FUNCTION_BLOCK Agua_Reuso (* Agua de reuso (serie 1000) - HidrycoLib *)
  (* Standard: 61499-2 *)
  (* Version 1.3, 20/10/2026, Hidryco, Hidryco, 1.3: simbolo sBoiaL (boia animada, verde/vermelho/cinza sem comunicacao). 1.2: o MGE do PCM Agua Reuso (MGE_1000) sai do CAT: passa a ser a instancia MGE_AGUA_REUSO do frame de MGEs do ETE_TJ; saem as saidas e tags do MGE. 1.1: MGE_1000 passa a ser o MGE_Generico (PM5300 pelo HW CAT PM53xxMbtcp, falta de fase e H/L de tensao e corrente); saidas stsFaltaFaseMGE, stsAlarmeMGE e stsPotenciaAtivaMGE; sai o cfgMonitoraMGE e o symlink stsConexaoMGE. 1.0: agua de reuso (serie 1000), so monitoracao. 1000-PIT-01/02 (Sensor_Generico, 4-20 mA, nivel) pelos symlinks ${PATH}PIT_1000_0x.stsSensorBruto; boia 1000-LSL-01 por ${PATH}stsBoiaLSL; comunicacao por ${PATH}stsFalhaRemota1 (BOOL, cartao), ${PATH}stsConexaoRemota2 e ${PATH}stsConexaoMGE (INT, connStatusInt); MGE do PCM Agua Reuso no MGE_1000. Valores e alarmes nas saidas do CAT. *)
  PACKAGE Hidryco.HidrycoLib;
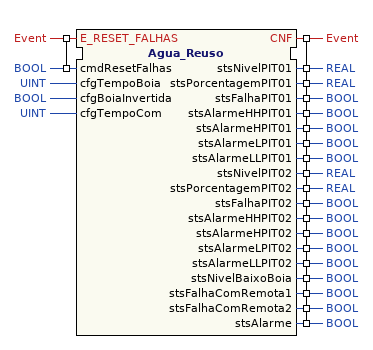
  EVENT_INPUT
    E_RESET_FALHAS WITH cmdResetFalhas; (* Reset pelo processo (sensores) com cmdResetFalhas = TRUE *)
  END_EVENT
  EVENT_OUTPUT
    CNF WITH stsNivelPIT01, stsPorcentagemPIT01, stsFalhaPIT01, stsAlarmeHHPIT01, stsAlarmeHPIT01, stsAlarmeLPIT01, stsAlarmeLLPIT01, stsNivelPIT02, stsPorcentagemPIT02, stsFalhaPIT02, stsAlarmeHHPIT02, stsAlarmeHPIT02, stsAlarmeLPIT02, stsAlarmeLLPIT02, stsNivelBaixoBoia, stsFalhaComRemota1, stsFalhaComRemota2, stsAlarme; (* Valores e alarmes (so na mudanca) *)
  END_EVENT
  VAR_INPUT
    cmdResetFalhas : BOOL; (* TRUE = reset (com o evento E_RESET_FALHAS) *)
    cfgTempoBoia : UINT := 10; (* Tempo (s) da boia 1000-LSL-01 abaixada para confirmar o nivel baixo *)
    cfgBoiaInvertida : BOOL := FALSE; (* FALSE: entrada da boia TRUE = nivel normal (boia levantada). TRUE: entrada TRUE = nivel baixo *)
    cfgTempoCom : UINT := 5; (* Tempo (s) sem comunicacao para confirmar a falha das remotas *)
  END_VAR
  VAR_OUTPUT
    stsNivelPIT01 : REAL; (* Nivel PIT_1000_01 (unidade de engenharia do sensor; 0 com o sinal em falha) *)
    stsPorcentagemPIT01 : REAL; (* Nivel PIT_1000_01 em % da altura maxima *)
    stsFalhaPIT01 : BOOL; (* Falha do sensor PIT_1000_01 (memorizada ate o reset) *)
    stsAlarmeHHPIT01 : BOOL; (* Alarme HH do PIT_1000_01 *)
    stsAlarmeHPIT01 : BOOL; (* Alarme H do PIT_1000_01 *)
    stsAlarmeLPIT01 : BOOL; (* Alarme L do PIT_1000_01 *)
    stsAlarmeLLPIT01 : BOOL; (* Alarme LL do PIT_1000_01 *)
    stsNivelPIT02 : REAL; (* Nivel PIT_1000_02 (unidade de engenharia do sensor; 0 com o sinal em falha) *)
    stsPorcentagemPIT02 : REAL; (* Nivel PIT_1000_02 em % da altura maxima *)
    stsFalhaPIT02 : BOOL; (* Falha do sensor PIT_1000_02 (memorizada ate o reset) *)
    stsAlarmeHHPIT02 : BOOL; (* Alarme HH do PIT_1000_02 *)
    stsAlarmeHPIT02 : BOOL; (* Alarme H do PIT_1000_02 *)
    stsAlarmeLPIT02 : BOOL; (* Alarme L do PIT_1000_02 *)
    stsAlarmeLLPIT02 : BOOL; (* Alarme LL do PIT_1000_02 *)
    stsNivelBaixoBoia : BOOL; (* Nivel baixo pela boia 1000-LSL-01 (confirmado por cfgTempoBoia) *)
    stsFalhaComRemota1 : BOOL; (* Falha de comunicacao com a remota 1 da Subestacao (boia) *)
    stsFalhaComRemota2 : BOOL; (* Falha de comunicacao com a remota 2 da Subestacao (PIT-01/02) *)
    stsAlarme : BOOL; (* Algum alarme da agua de reuso (sensores, boia, comunicacao) *)
  END_VAR
  FBS
    IThis : Agua_Reuso_HMI(QI := TRUE);
    plcStart1 : plcStart(Prio := 10);
    Logica : basicAguaReuso;
    Tick : E_CYCLE(DT := T#1s);
    PIT_1000_01 : Sensor_Generico(pin_FC98F78ABCBC0A7E := TRUE, pin_CC8EEC06FF0C4430 := 'm', pin_D46B37D45FD5AF5D := FALSE, pin_31E57DCE3AF9C996 := 4000.0, pin_BFED79817B71957D := 20000.0, pin_CA39953142B1EBBD := 3800.0, pin_519A2B73CC673344 := 22000.0, pin_F21E4E6BC95CB4D0 := 5, pin_0ECE7B3867B02E0B := FALSE, pin_6D3A2524C5D0F0D1 := 2);
    PIT_1000_02 : Sensor_Generico(pin_FC98F78ABCBC0A7E := TRUE, pin_CC8EEC06FF0C4430 := 'm', pin_D46B37D45FD5AF5D := FALSE, pin_31E57DCE3AF9C996 := 4000.0, pin_BFED79817B71957D := 20000.0, pin_CA39953142B1EBBD := 3800.0, pin_519A2B73CC673344 := 22000.0, pin_F21E4E6BC95CB4D0 := 5, pin_0ECE7B3867B02E0B := FALSE, pin_6D3A2524C5D0F0D1 := 2);
    BoiaLSL : SYMLINKMULTIVARDST_1559B0FF8170C9BA0(NAME1 := '$${PATH}stsBoiaLSL', QI := TRUE); {SET_ATTRIBUTE(Configuration.GenericFBType.InterfaceParams, Runtime.System#I:=1;VALUE${I$}:BOOL)}
    FalhaRemota1 : SYMLINKMULTIVARDST_1559B0FF8170C9BA0(NAME1 := '$${PATH}stsFalhaRemota1', QI := TRUE); {SET_ATTRIBUTE(Configuration.GenericFBType.InterfaceParams, Runtime.System#I:=1;VALUE${I$}:BOOL)}
    ConexaoRemota2 : SYMLINKMULTIVARDST_5A03F112CD5D470(NAME1 := '$${PATH}stsConexaoRemota2', QI := TRUE); {SET_ATTRIBUTE(Configuration.GenericFBType.InterfaceParams, Runtime.System#I:=1;VALUE${I$}:INT)}
    AlarmeNivelBaixo : ALARM_BIT(TYPE := 1, ACKTYPE_1 := 2, ACTIVE := TRUE); {SET_ATTRIBUTE(HMI.AlarmText, Nível baixo no reservatório (boia 1000-LSL-01))} {SET_ATTRIBUTE(HMI.AlarmClass, Warning)}
    AlarmeRemota1 : ALARM_BIT(TYPE := 1, ACKTYPE_1 := 2, ACTIVE := TRUE); {SET_ATTRIBUTE(HMI.AlarmText, Remota 1 da Subestação sem comunicação (boia 1000-LSL-01))}
    AlarmeRemota2 : ALARM_BIT(TYPE := 1, ACKTYPE_1 := 2, ACTIVE := TRUE); {SET_ATTRIBUTE(HMI.AlarmText, Remota 2 da Subestação sem comunicação (1000-PIT-01/02))}
  END_FBS
  EVENT_CONNECTIONS
    plcStart1.FIRST_INIT TO IThis.5B291D4D67D48173;
    plcStart1.REDO_INIT TO IThis.5B291D4D67D48173;
    IThis.D656758D65B70390 TO Logica.1F2574A6F30133E3;
    Logica.82CEBA2D0471C377 TO Tick.START;
    Logica.82CEBA2D0471C377 TO BoiaLSL.INIT;
    Logica.82CEBA2D0471C377 TO FalhaRemota1.INIT;
    Logica.82CEBA2D0471C377 TO ConexaoRemota2.INIT;
    Logica.82CEBA2D0471C377 TO AlarmeNivelBaixo.INIT;
    AlarmeNivelBaixo.INITO TO AlarmeNivelBaixo.REQ_INITDATA;
    AlarmeNivelBaixo.CNF_INITDATA TO AlarmeNivelBaixo.ACTIVATE;
    AlarmeNivelBaixo.INITO TO AlarmeRemota1.INIT;
    AlarmeRemota1.INITO TO AlarmeRemota1.REQ_INITDATA;
    AlarmeRemota1.CNF_INITDATA TO AlarmeRemota1.ACTIVATE;
    AlarmeRemota1.INITO TO AlarmeRemota2.INIT;
    AlarmeRemota2.INITO TO AlarmeRemota2.REQ_INITDATA;
    AlarmeRemota2.CNF_INITDATA TO AlarmeRemota2.ACTIVATE;
    AlarmeRemota2.INITO TO plcStart1.ACK_FIRST;
    AlarmeRemota2.INITO TO IThis.BA9200524709281B;
    IThis.05D27B56DB642E3B TO Logica.196CC39C90BB2858;
    E_RESET_FALHAS TO Logica.F8A99F29850AD5DB;
    BoiaLSL.CNF TO Logica.299D414224484D8E;
    FalhaRemota1.CNF TO Logica.AF9BA5F5EA0D0DE5;
    ConexaoRemota2.CNF TO Logica.AF9BA5F5EA0D0DE5;
    Tick.EO TO Logica.FD7FC9E3C7412179;
    Logica.0D7078056D047821 TO CNF;
    Logica.48B7766158A72DB1 TO IThis.0FFD476B12261BFC;
    PIT_1000_01.28A380156DB271B8 TO Logica.B449598857AB2011;
    Logica.D611B8DF03491A62 TO PIT_1000_01.D21DAA5004F58516;
    PIT_1000_02.28A380156DB271B8 TO Logica.25FCE411FF203199;
    Logica.D611B8DF03491A62 TO PIT_1000_02.D21DAA5004F58516;
    Logica.A53CD1FF4E04D581 TO AlarmeNivelBaixo.REQ;
    Logica.A53CD1FF4E04D581 TO AlarmeRemota1.REQ;
    Logica.A53CD1FF4E04D581 TO AlarmeRemota2.REQ;
    AlarmeNivelBaixo.IND_1 TO IThis.0FFD476B12261BFC;
    AlarmeRemota1.IND_1 TO IThis.0FFD476B12261BFC;
    AlarmeRemota2.IND_1 TO IThis.0FFD476B12261BFC;
    IThis.05D27B56DB642E3B TO AlarmeNivelBaixo.ACK_C1;
    IThis.05D27B56DB642E3B TO AlarmeRemota1.ACK_C1;
    IThis.05D27B56DB642E3B TO AlarmeRemota2.ACK_C1;
  END_CONNECTIONS
  DATA_CONNECTIONS
    cfgTempoBoia TO Logica.7AB282FA59C5DE18;
    cfgBoiaInvertida TO Logica.78056A861A9FC565;
    cfgTempoCom TO Logica.DDE31F23C75A7867;
    cmdResetFalhas TO Logica.4012098E9C8C3E1C;
    PIT_1000_01.D7422D307E6AF52D TO Logica.07D3FD1B9693EBA9;
    PIT_1000_01.E6F78A591442B69F TO Logica.1ED47B1DA7FFFE36;
    PIT_1000_01.07C3588C57A022B8 TO Logica.4674F0A0B1306602;
    PIT_1000_01.726640D1704B3F86 TO Logica.483E654AA9295F1F;
    PIT_1000_01.6108F9B5CA5170A6 TO Logica.2F7955EE24BC434E;
    PIT_1000_01.9578190A49DBC450 TO Logica.AFE2694C114D5BB0;
    PIT_1000_01.0D14BA934DBED883 TO Logica.586B59BB34B41275;
    PIT_1000_01.ADAD629D7A214F32 TO Logica.F32A97D9BEF784AF;
    PIT_1000_01.53279A5859ECAB18 TO Logica.A3BCA6E4A914D759;
    Logica.E0009B8BCCB1DC9C TO PIT_1000_01.1908F43CB878F5E7;
    PIT_1000_02.D7422D307E6AF52D TO Logica.D111AE3CF546FB41;
    PIT_1000_02.E6F78A591442B69F TO Logica.538692287664FC27;
    PIT_1000_02.07C3588C57A022B8 TO Logica.67FA77966B860F92;
    PIT_1000_02.726640D1704B3F86 TO Logica.785FA5DCD1BD1BBE;
    PIT_1000_02.6108F9B5CA5170A6 TO Logica.129365CAD32FA68D;
    PIT_1000_02.9578190A49DBC450 TO Logica.768E3A7133E77018;
    PIT_1000_02.0D14BA934DBED883 TO Logica.834EF20FB7F0A45B;
    PIT_1000_02.ADAD629D7A214F32 TO Logica.AD38A0A4A9FD5CE4;
    PIT_1000_02.53279A5859ECAB18 TO Logica.2BF6430062E3707F;
    Logica.E0009B8BCCB1DC9C TO PIT_1000_02.1908F43CB878F5E7;
    BoiaLSL.VALUE1 TO Logica.B38FC6C6C258CD1C;
    FalhaRemota1.VALUE1 TO Logica.E3D9D2003045C208;
    ConexaoRemota2.VALUE1 TO Logica.9A84D5DA142F5D34;
    IThis.8080CCD0B707ACBC TO Logica.A39AEE8EBC0FF16A;
    Logica.06A990B615DC7EBF TO AlarmeNivelBaixo.INP;
    Logica.8FB5C28302258408 TO AlarmeRemota1.INP;
    Logica.45C3A871E8411D0B TO AlarmeRemota2.INP;
    Logica.CA2E43CC2AB7A710 TO stsNivelPIT01;
    Logica.EFF4A50248596AAE TO stsPorcentagemPIT01;
    Logica.D29D6389261AB801 TO stsFalhaPIT01;
    Logica.C356053499FD22FD TO stsAlarmeHHPIT01;
    Logica.6D07A7E00D0B552D TO stsAlarmeHPIT01;
    Logica.E662ECFBF9CE0E97 TO stsAlarmeLPIT01;
    Logica.DAE46A0ED33EAB6E TO stsAlarmeLLPIT01;
    Logica.68F5A0DB478BBF75 TO stsNivelPIT02;
    Logica.38F9A56D3A39F26B TO stsPorcentagemPIT02;
    Logica.C6322136FABA67B7 TO stsFalhaPIT02;
    Logica.25F036F3521BEB36 TO stsAlarmeHHPIT02;
    Logica.DCDA1244C5EBD289 TO stsAlarmeHPIT02;
    Logica.AC8C91AE55FF19B5 TO stsAlarmeLPIT02;
    Logica.CE4E9CC28966EAEA TO stsAlarmeLLPIT02;
    Logica.02BA5107AB682069 TO stsNivelBaixoBoia;
    Logica.E4841A579A62D291 TO stsFalhaComRemota1;
    Logica.737542A8C4F021EE TO stsFalhaComRemota2;
    Logica.6565994057372119 TO stsAlarme;
    Logica.CA2E43CC2AB7A710 TO IThis.502DB12634FA3EAE;
    Logica.EFF4A50248596AAE TO IThis.81C0628EFE8726A6;
    Logica.6F6AFBBD21CDC2A9 TO IThis.35A08BB1DE44C71A;
    Logica.68F5A0DB478BBF75 TO IThis.A8D89D8718373A64;
    Logica.38F9A56D3A39F26B TO IThis.2529D64949E9AEE6;
    Logica.D04BD5C366CB1C25 TO IThis.E2AEEC2ED3B0FA82;
    Logica.3319F6072649D6C8 TO IThis.C99A868607210194;
    Logica.02BA5107AB682069 TO IThis.F60000E1A4383811;
    Logica.E4841A579A62D291 TO IThis.BF5934575D19358B;
    Logica.737542A8C4F021EE TO IThis.87D3EF366AF9B5C3;
    Logica.6565994057372119 TO IThis.759FEBA1D038B19B;
    AlarmeNivelBaixo.STATE_1 TO IThis.1946141CF0DDF720;
    AlarmeRemota1.STATE_1 TO IThis.B090B8451459FC56;
    AlarmeRemota2.STATE_1 TO IThis.FB7C34D2BA98C96C;
  END_CONNECTIONS
END_FUNCTION_BLOCK
